{region 'Documentation'}
(*!
<summary>Check that IN is at most Maximum.</summary>
*)
{endregion}
FUNCTION_BLOCK AssertLessEqual_UInt EXTENDS AssertionBase
VAR_INPUT
    IN : UINT; //! Actual value checked or observed by this Assertion.
    Maximum : UINT; //! Inclusive upper bound of the comparison; for a range, must not be below Minimum.
END_VAR

SUPER^();

{region 'Documentation'}
(*!
<summary>Check that IN is at most Maximum.</summary>
*)
{endregion}
METHOD PROTECTED Assert
VAR
    Message : STRING(GVL_Constants.MessageLength);
    MaximumText : STRING(GVL_Constants.AssertionValueLength);
    ActualText : STRING(GVL_Constants.AssertionValueLength);
END_VAR
IF NOT EvaluationActive THEN
    RETURN;
END_IF;

IF Result = E_Result.Error THEN
    RETURN;
END_IF;

IF Result = E_Result.Failed THEN
    RETURN;
END_IF;

IF IN > Maximum THEN
    MaximumText := UINT_TO_STRING(Maximum);
    ActualText := UINT_TO_STRING(IN);
    Message := CONCAT('Assertion failed: value is above maximum. Maximum = ',
        MaximumText);
    Message := CONCAT(Message, ', Actual = ');
    Message := CONCAT(Message, ActualText);
    Message := CONCAT(Message, '.');
    Fail(Message := Message);
    RETURN;
END_IF;

Pass();
END_METHOD

END_FUNCTION_BLOCK

(* stored: Version 1.1.0.1
   POU AssertLessEqual_UInt: Id {1dc46eef-af3d-4120-bc39-f7b8bedb78b2}, SpecialFunc None
   Folder Internal: Id {1ffff991-eee5-47f7-a08c-ea3ea1d4e987}
   Method Assert: Id {cd6daacd-120f-403c-8adf-4bddc88c6e64} *)
